{attribute 'qualified_only'}
{attribute 'strict'}
{attribute 'to_string'}
TYPE E_SeverityNumber :
(
	UNSPECIFIED := 0,
	TRACE,
	TRACE2,
	TRACE3,
	TRACE4,
	DEBUG,
	DEBUG2,
	DEBUG3,
	DEBUG4,
	INFO,
	INFO2,
	INFO3,
	INFO4,
	WARN,
	WARN2,
	WARN3,
	WARN4,
	ERROR,
	ERROR2,
	ERROR3,
	ERROR4,
	FATAL,
	FATAL2,
	FATAL3,
	FATAL4
);
END_TYPE

(* stored: Version 1.1.0.1
   EnumerationTextList E_SeverityNumber: Id {42fbc878-be73-47d8-84c4-df1caec01f70} *)
